TEXTLIST TextList_Piston_Recipe_State_InOut
  0 = ' '
  1 = 'In'
  2 = 'Out'
   = ''
END_TEXTLIST

(* stored: Version 1.1.0.1, ProductVersion 3.1.4024.12
   TextList TextList_Piston_Recipe_State_InOut: Id {5cb0fdc2-f5be-43ae-902a-ace45a36aa40} *)
